FUNCTION F_TimeRatio : INT
VAR_INPUT
	t1: TIME;
	t2: TIME;

END_VAR
VAR
	udi_t1: UDINT;
	udi_t2: UDINT;

	ratio: REAL;
END_VAR


udi_t1:=TIME_TO_UDINT(t1);
udi_t2:=TIME_TO_UDINT(t2);

IF udi_t2>0 THEN;
	ratio:=udi_t1/udi_t2;
END_IF

END_FUNCTION

(* stored: Version 1.1.0.1, ProductVersion 3.1.4024.12
   POU F_TimeRatio: Id {9e63d04d-22ba-44b7-a7dd-32366321d33f}, SpecialFunc None *)
